(*
SPDX-FileCopyrightText: © 2026 Oleksandr Tiutyk <trofimich@gmail.com>
SPDX-License-Identifier: MIT
License: https://opensource.org/license/mit
*)

(*!
<summary>
Beckhoff EL3413: 3-phase power measurement terminal up to 690 V AC.
</summary>
<description>
Represents phase TxPDOs 0x1A00..0x1A02, auxiliary TxPDO 0x1A03,
phase selector RxPDOs 0x1600..0x1602 and auxiliary selector RxPDO 0x1603.
Phase and auxiliary Status fields are required; bit 14 invalidates the corresponding measurement.
Bus WcState and State do not replace measurement status. Interpret values using acknowledged input selectors.
Units and additional index selections follow firmware and configured transformer ratios.
Link fields individually. Use one owner task and synchronize other access; snapshots are not atomic.
When used for I/O, link located fields or their containing buffers to the matching selected PDOs.
The record is not a packed wire buffer; compiler padding is not part of the device specification.
Unlinked/default values do not prove valid I/O. The caller evaluates bus/channel validity before use.
Use one owner task per instance and externally synchronize other access; multi-field snapshots are not atomic.
Copies store data without creating hardware links. Keep borrowed field references valid while consumers are bound.
This passive record performs no validation, synchronization, configuration or protocol advancement.
</description>
*)
TYPE EL3413 :
STRUCT
	L1 : POWER_MEASUREMENT_CHANNEL;
	L2 : POWER_MEASUREMENT_CHANNEL;
	L3 : POWER_MEASUREMENT_CHANNEL;
	Auxiliary : POWER_MEASUREMENT_AUXILIARY_CHANNEL;
END_STRUCT
END_TYPE

(* stored: Version 1.1.0.1, ProductVersion 3.1.4026.20
   DUT EL3413: Id {6c58d245-21ab-4b92-bb4f-1b6cf5dffe0d} *)
